// TIA Portal V21 export
// export: Created 2026-10-12T11:32:15.8965028Z, ExportSetting WithDefaults, DisplayName Totally Integrated Automation Portal, DisplayVersion V21, DisplayName STEP 7 Professional, DisplayVersion V21, DisplayName STEP 7 Safety, DisplayVersion V21, DisplayName Tech WebApplication, DisplayVersion V21, DisplayName WinCC Basic/Comfort/Advanced, DisplayVersion V21, DisplayName WinCC Unified, DisplayVersion V21
FUNCTION "FC_AUTO" : Void   // FC5, LAD
{ S7_Optimized_Access := 'TRUE' }
VERSION : 0.1
// stored: AutoNumber true, IsIECCheckEnabled false, SetENOAutomatically false, UDAEnableTagReadback false
   VAR_TEMP   // added for the SCL form of the ladder/FBD networks
      _w1 : Bool;
      _w2 : Bool;
      _w3 : Bool;
   END_VAR
BEGIN

REGION Network 1: AUTO ON
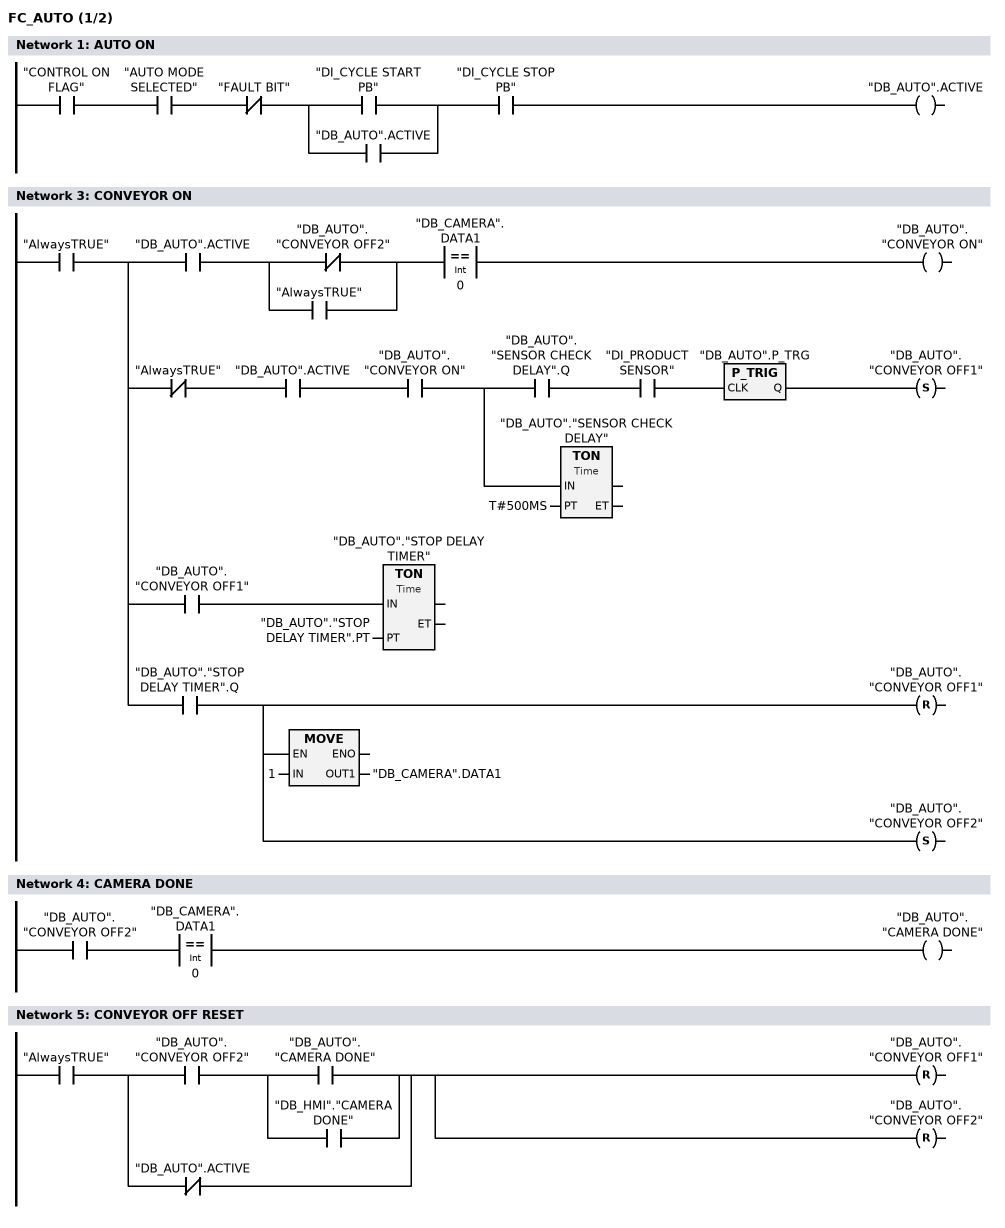
   RUNG wire#powerrail
      Contact( "CONTROL ON FLAG" )
      Contact( "AUTO MODE SELECTED" )
      I_Contact( "FAULT BIT" )
      wire#w1
      Contact( "DI_CYCLE START PB" )
      wire#w2
      Contact( "DI_CYCLE STOP PB" )
      Coil( "DB_AUTO".ACTIVE )
   END_RUNG
   RUNG wire#w1
      Contact( "DB_AUTO".ACTIVE )
   END_RUNG wire#w2
   // the same network as SCL:
   "DB_AUTO".ACTIVE := "CONTROL ON FLAG" AND "AUTO MODE SELECTED" AND NOT "FAULT BIT" AND ("DI_CYCLE START PB" OR "DB_AUTO".ACTIVE) AND "DI_CYCLE STOP PB";
END_REGION

REGION Network 2 (SCL): STOP DELAY TIME
   "DB_AUTO"."STOP DELAY TIMER".PT := "DB_HMI"."STOP TIME" * 1000;
END_REGION

REGION Network 3: CONVEYOR ON
   RUNG wire#powerrail
      Contact( "AlwaysTRUE" )
      wire#w1
      Contact( "DB_AUTO".ACTIVE )
      wire#w2
      I_Contact( "DB_AUTO"."CONVEYOR OFF2" )
      wire#w3
      { S7_Templates := "SrcType := Int" } EQ_Contact(in1 := "DB_CAMERA".DATA1, in2 := 0)
      Coil( "DB_AUTO"."CONVEYOR ON" )
   END_RUNG
   RUNG wire#w2
      Contact( "AlwaysTRUE" )
   END_RUNG wire#w3
   RUNG wire#w1
      I_Contact( "AlwaysTRUE" )
      Contact( "DB_AUTO".ACTIVE )
      Contact( "DB_AUTO"."CONVEYOR ON" )
      wire#w4
      Contact( "DB_AUTO"."SENSOR CHECK DELAY".Q )
      Contact( "DI_PRODUCT SENSOR" )
      P_Trig( "DB_AUTO".P_TRG )
      S_Coil( "DB_AUTO"."CONVEYOR OFF1" )
   END_RUNG
   RUNG wire#w4
      { S7_Templates := "time_type := Time" } "DB_AUTO"."SENSOR CHECK DELAY".TON(pt := T#500MS, et =>)
   END_RUNG
   RUNG wire#w1
      Contact( "DB_AUTO"."CONVEYOR OFF1" )
      { S7_Templates := "time_type := Time" } "DB_AUTO"."STOP DELAY TIMER".TON(pt := "DB_AUTO"."STOP DELAY TIMER".PT, et =>)
   END_RUNG
   RUNG wire#w1
      Contact( "DB_AUTO"."STOP DELAY TIMER".Q )
      wire#w5
      R_Coil( "DB_AUTO"."CONVEYOR OFF1" )
   END_RUNG
   RUNG wire#w5
      Move(in := 1, out1 => "DB_CAMERA".DATA1)
   END_RUNG
   RUNG wire#w5
      S_Coil( "DB_AUTO"."CONVEYOR OFF2" )
   END_RUNG
   // the same network as SCL:
   "DB_AUTO"."CONVEYOR ON" := "AlwaysTRUE" AND "DB_AUTO".ACTIVE AND (NOT "DB_AUTO"."CONVEYOR OFF2" OR "AlwaysTRUE") AND ("DB_CAMERA".DATA1 = 0);
   #_w1 := "AlwaysTRUE" AND NOT "AlwaysTRUE" AND "DB_AUTO".ACTIVE AND "DB_AUTO"."CONVEYOR ON";
   #_w2 := #_w1 AND "DB_AUTO"."SENSOR CHECK DELAY".Q AND "DI_PRODUCT SENSOR";
   #_w3 := #_w2 AND NOT "DB_AUTO".P_TRG;   // rising edge
   "DB_AUTO".P_TRG := #_w2;
   IF #_w3 THEN "DB_AUTO"."CONVEYOR OFF1" := TRUE; END_IF;
   "DB_AUTO"."SENSOR CHECK DELAY".TON(IN := #_w1, PT := T#500MS);
   "DB_AUTO"."STOP DELAY TIMER".TON(IN := "AlwaysTRUE" AND "DB_AUTO"."CONVEYOR OFF1",
                           PT := "DB_AUTO"."STOP DELAY TIMER".PT);
   IF "AlwaysTRUE" AND "DB_AUTO"."STOP DELAY TIMER".Q THEN
       "DB_AUTO"."CONVEYOR OFF1" := FALSE;
       "DB_CAMERA".DATA1 := 1;
       "DB_AUTO"."CONVEYOR OFF2" := TRUE;
   END_IF;
END_REGION

REGION Network 4: CAMERA DONE
   RUNG wire#powerrail
      Contact( "DB_AUTO"."CONVEYOR OFF2" )
      { S7_Templates := "SrcType := Int" } EQ_Contact(in1 := "DB_CAMERA".DATA1, in2 := 0)
      Coil( "DB_AUTO"."CAMERA DONE" )
   END_RUNG
   // the same network as SCL:
   "DB_AUTO"."CAMERA DONE" := "DB_AUTO"."CONVEYOR OFF2" AND ("DB_CAMERA".DATA1 = 0);
END_REGION

REGION Network 5: CONVEYOR OFF RESET
   RUNG wire#powerrail
      Contact( "AlwaysTRUE" )
      wire#w1
      Contact( "DB_AUTO"."CONVEYOR OFF2" )
      wire#w2
      Contact( "DB_AUTO"."CAMERA DONE" )
      wire#w3
      R_Coil( "DB_AUTO"."CONVEYOR OFF1" )
   END_RUNG
   RUNG wire#w2
      Contact( "DB_HMI"."CAMERA DONE" )
   END_RUNG wire#w3
   RUNG wire#w1
      I_Contact( "DB_AUTO".ACTIVE )
   END_RUNG wire#w3
   RUNG wire#w3
      R_Coil( "DB_AUTO"."CONVEYOR OFF2" )
   END_RUNG
   // the same network as SCL:
   IF "AlwaysTRUE" AND (("DB_AUTO"."CONVEYOR OFF2" AND ("DB_AUTO"."CAMERA DONE" OR "DB_HMI"."CAMERA DONE")) OR NOT "DB_AUTO".ACTIVE) THEN
       "DB_AUTO"."CONVEYOR OFF1" := FALSE;
       "DB_AUTO"."CONVEYOR OFF2" := FALSE;
   END_IF;
END_REGION

REGION Network 6: AUTO STATUS
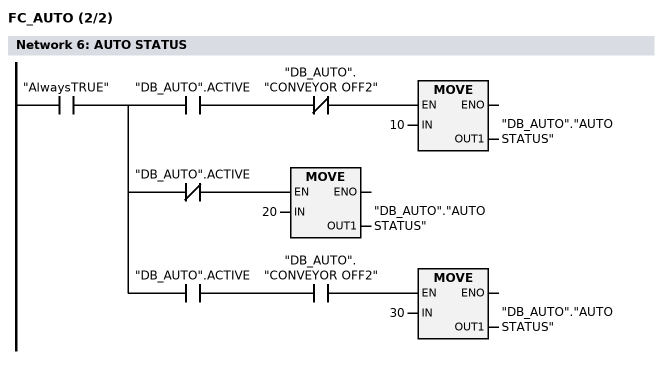
   RUNG wire#powerrail
      Contact( "AlwaysTRUE" )
      wire#w1
      Contact( "DB_AUTO".ACTIVE )
      I_Contact( "DB_AUTO"."CONVEYOR OFF2" )
      Move(in := 10, out1 => "DB_AUTO"."AUTO STATUS")
   END_RUNG
   RUNG wire#w1
      I_Contact( "DB_AUTO".ACTIVE )
      Move(in := 20, out1 => "DB_AUTO"."AUTO STATUS")
   END_RUNG
   RUNG wire#w1
      Contact( "DB_AUTO".ACTIVE )
      Contact( "DB_AUTO"."CONVEYOR OFF2" )
      Move(in := 30, out1 => "DB_AUTO"."AUTO STATUS")
   END_RUNG
   // the same network as SCL:
   IF "AlwaysTRUE" AND "DB_AUTO".ACTIVE AND NOT "DB_AUTO"."CONVEYOR OFF2" THEN
       "DB_AUTO"."AUTO STATUS" := 10;
   END_IF;
   IF "AlwaysTRUE" AND NOT "DB_AUTO".ACTIVE THEN "DB_AUTO"."AUTO STATUS" := 20; END_IF;
   IF "AlwaysTRUE" AND "DB_AUTO".ACTIVE AND "DB_AUTO"."CONVEYOR OFF2" THEN
       "DB_AUTO"."AUTO STATUS" := 30;
   END_IF;
END_REGION
END_FUNCTION
